(* IEC 61131-3 sources: trust-platform/examples/control/01-feedback-foundations-and-temperature-control/08-heating-valve-rate-tracking/src, 2 files *)

(* ---- Main.st ---- *)
USING Control;

(* Fraction of the raw-minus-filtered difference applied per update: alpha = dt/(Tf + dt). *)
FUNCTION FilterFraction : LREAL
VAR_INPUT
    CycleTime : LREAL;
    FilterTime : LREAL;
END_VAR
FilterFraction := CycleTime / (FilterTime + CycleTime);
END_FUNCTION

(* First-order low-pass update: yf_new = yf_old + alpha·(yr − yf_old). *)
FUNCTION FilterUpdate : LREAL
VAR_INPUT
    PreviousFilteredValue : LREAL;
    RawValue : LREAL;
    FilterFraction : LREAL;
END_VAR
FilterUpdate := PreviousFilteredValue + FilterFraction * (RawValue - PreviousFilteredValue);
END_FUNCTION

(* An interval is usable only if time has advanced and the samples can still represent the
   loop's fastest oscillation. *)
FUNCTION IntervalUsable : BOOL
VAR_INPUT
    ElapsedTime : LREAL;
    MaximumInterval : LREAL;
END_VAR
IntervalUsable := ElapsedTime > LREAL#0.0 AND ElapsedTime <= MaximumInterval;
END_FUNCTION

(* Integral correction toward the measured actuator position: I_next = I* + dt/Tt·(x − u_r). *)
FUNCTION MeasuredTrackingCorrection : LREAL
VAR_INPUT
    StemPosition : LREAL;
    Request : LREAL;
    Elapsed : LREAL;
    TrackingTime : LREAL;
END_VAR
MeasuredTrackingCorrection := Elapsed / TrackingTime * (StemPosition - Request);
END_FUNCTION

(* A reading is usable only with good source quality, inside the sensor's 0–80 °C range and with an age
   between 0 and MaximumAge. NaN fails every comparison. *)
FUNCTION ReadingUsable : BOOL
VAR_INPUT
    QualityGood : BOOL;
    Value : LREAL;
    Age : LREAL;
    MaximumAge : LREAL;
END_VAR
ReadingUsable := QualityGood AND Value >= LREAL#0.0 AND Value <= LREAL#80.0
    AND Age >= LREAL#0.0 AND Age <= MaximumAge;
END_FUNCTION

(* Weighted proportional term about the operating point T0: P = Kp·(β·(SP − T0) − (PV − T0)). *)
FUNCTION WeightedProportional : LREAL
VAR_INPUT
    ProportionalGain : LREAL;
    SetpointWeight : LREAL;
    Setpoint : LREAL;
    ProcessValue : LREAL;
    OperatingPoint : LREAL;
END_VAR
WeightedProportional := ProportionalGain
    * (SetpointWeight * (Setpoint - OperatingPoint) - (ProcessValue - OperatingPoint));
END_FUNCTION

(* Integral state that makes P + I reproduce the applied command: I = u_applied − P. *)
FUNCTION InitialIntegral : LREAL
VAR_INPUT
    AppliedOutput : LREAL;
    Proportional : LREAL;
END_VAR
InitialIntegral := AppliedOutput - Proportional;
END_FUNCTION

(* A candidate set is usable only as a whole: non-negative gains, weights in 0–1, a minimum below the
   maximum, rate limits around zero, a positive tracking time and a non-negative filter time.
   Any NaN fails its comparison and rejects the set. *)
FUNCTION ValidPidParameters : BOOL
VAR_INPUT
    Candidate : Control.PIDParameters;
    FilterTime : LREAL;
END_VAR
ValidPidParameters :=
    Candidate.ProportionalGain >= LREAL#0.0 AND Candidate.IntegralGain >= LREAL#0.0
    AND Candidate.DerivativeGain >= LREAL#0.0
    AND Candidate.ProportionalSetpointWeight >= LREAL#0.0 AND Candidate.ProportionalSetpointWeight <= LREAL#1.0
    AND Candidate.DerivativeSetpointWeight >= LREAL#0.0 AND Candidate.DerivativeSetpointWeight <= LREAL#1.0
    AND Candidate.Bias = Candidate.Bias
    AND Candidate.OutputMinimum < Candidate.OutputMaximum
    AND Candidate.RateMinimum <= LREAL#0.0 AND Candidate.RateMaximum >= LREAL#0.0
    AND Candidate.TrackingTime > LREAL#0.0
    AND FilterTime >= LREAL#0.0;
END_FUNCTION

FUNCTION SamePidParameters : BOOL
VAR_INPUT
    Left : Control.PIDParameters;
    Right : Control.PIDParameters;
END_VAR
SamePidParameters :=
    Left.ProportionalGain = Right.ProportionalGain
    AND Left.IntegralGain = Right.IntegralGain
    AND Left.DerivativeGain = Right.DerivativeGain
    AND Left.ProportionalSetpointWeight = Right.ProportionalSetpointWeight
    AND Left.DerivativeSetpointWeight = Right.DerivativeSetpointWeight
    AND Left.Bias = Right.Bias
    AND Left.OutputMinimum = Right.OutputMinimum
    AND Left.OutputMaximum = Right.OutputMaximum
    AND Left.RateMinimum = Right.RateMinimum
    AND Left.RateMaximum = Right.RateMaximum
    AND Left.TrackingTime = Right.TrackingTime
    AND Left.AntiWindup = Right.AntiWindup;
END_FUNCTION

PROGRAM Main
VAR
    Controller : Control.PID;
    (* Tune replaces this record with each candidate; the defaults are the controller commissioned
       on the electric heater in Lesson 30. *)
    Parameters : Control.PIDParameters := (
        ProportionalGain := LREAL#13.0,
        IntegralGain := LREAL#3.5,
        DerivativeGain := LREAL#0.0,
        ProportionalSetpointWeight := LREAL#0.3,
        DerivativeSetpointWeight := LREAL#0.0,
        Bias := LREAL#0.0,
        OutputMinimum := LREAL#0.0,
        OutputMaximum := LREAL#100.0,
        RateMinimum := LREAL#-10000.0,
        RateMaximum := LREAL#10000.0,
        TrackingTime := LREAL#1.0,
        AntiWindup := PIDAntiWindup#BackCalculation
    );
    ConfiguredParameters : Control.PIDParameters;
    ConfiguredFilterTimeS : LREAL := 1.0;
    ParameterRevision : DINT := 0;
    ParametersRejected : BOOL := FALSE;
    InitialState : Control.PIDInitialState;
    ObservedState : Control.PIDInitialState;
    Input : Control.PIDInput;
    (* Ready: every retained value has been set from the actual operating condition. *)
    Initialized : BOOL := FALSE;
    InitializeRequest : BOOL := FALSE;
    InitializeRequestWas : BOOL := FALSE;
    AutoMode : BOOL := FALSE;
    AutoActive : BOOL := FALSE;
    (* TRUE at start: a program that starts in Auto from preset stored values continues without a
       transfer. A real start begins uninitialized in Manual, which clears it. *)
    AutoWasActive : BOOL := TRUE;
    (* FALSE runs the untracked counterexample: Manual leaves the stored values as initialized. *)
    TrackManual : BOOL := TRUE;
    ManualOutput : LREAL := 75.0;
    (* Sensor interface: the simulated device delivers the reading with a quality flag; these three
       inputs inject faults for the lesson. *)
    SensorQualityGood : BOOL := TRUE;
    SensorFrozen : BOOL := FALSE;
    InjectedOffsetC : LREAL := 0.0;
    ReadingC : LREAL := 35.0;
    AcquisitionTimer : TON;
    AcquisitionAgeS : LREAL := 0.0;
    NewAcquisition : BOOL := FALSE;
    (* Measurement validity: a reading older than MaximumAgeS is stale; recovery needs
       FreshSamplesRequired consecutive fresh valid acquisitions after an acknowledgement. *)
    MaximumAgeS : LREAL := 0.5;
    FreshSamplesRequired : DINT := 3;
    MeasurementUsable : BOOL := FALSE;
    MeasurementFault : BOOL := FALSE;
    FaultAcknowledge : BOOL := FALSE;
    Acknowledged : BOOL := FALSE;
    RecoveryCount : DINT := 0;
    RecoveryComplete : BOOL := FALSE;
    SetpointC : LREAL := 35.0;
    TemperatureC : LREAL := 35.0;
    SafeProcessValueC : LREAL := 35.0;
    (* Requested position, bounded target and measured position: the PI request before the 0–100 %
       limits, the target sent to the valve, and the stem position the valve has reached. *)
    NominalRequestPct : LREAL := 75.0;
    ValveRequestPct : LREAL := 75.0;
    StemPositionPct : LREAL := 75.0;
    (* FALSE tracks only the bounded target: the counterexample. *)
    TrackMeasuredPosition : BOOL := TRUE;
    TrackingCorrectionPct : LREAL := 0.0;
    ErrorC : LREAL := 0.0;
    (* Reference of the weighted proportional term: the 35 °C hot operating point. *)
    OperatingPointC : LREAL := 35.0;
    (* Measurement filter: Tf = 0 bypasses it; Control Studio applies Tf with the gains. *)
    FilterTimeS : LREAL := 1.0;
    FilterAlpha : LREAL := 1.0;
    FilteredC : LREAL := 35.0;
    FilterRestart : BOOL := TRUE;
    (* Timing: the controller updates every ControllerPeriodS of measured time. *)
    IntervalTimer : TON;
    SinceLastUpdateS : LREAL := 0.0;
    ElapsedS : LREAL := 0.0;
    ControllerPeriodS : LREAL := 0.1;
    (* Longest usable interval: half the loop's 4.42 s ultimate period (Lesson 20). *)
    MaximumIntervalS : LREAL := 2.2;
    UpdateDue : BOOL := FALSE;
    TimingUsable : BOOL := FALSE;
    RejectedUpdates : DINT := 0;
    ProportionalPct : LREAL := 0.0;
    IntegralPct : LREAL := 75.0;
    PreviousRequestPct : LREAL := 75.0;
    CommandActivityPoints : LREAL := 0.0;
END_VAR

(* The water heated through the valve; the temperature measurement carries ±0.02 °C noise. *)
(* Sensor interface: every scan the device delivers a new acquisition unless it is frozen. The
   acquisition timer restarts with each new acquisition, so its elapsed time is the reading's age. *)
IF NOT SensorFrozen THEN
    ReadingC := TemperatureC + InjectedOffsetC;
    AcquisitionTimer(IN := FALSE, PT := T#1h);
    NewAcquisition := TRUE;
ELSE
    NewAcquisition := FALSE;
END_IF;
AcquisitionTimer(IN := TRUE, PT := T#1h);
AcquisitionAgeS := UDINT_TO_LREAL(DWORD_TO_UDINT(TIME_TO_DWORD(AcquisitionTimer.ET))) / LREAL#1000.0;

MeasurementUsable := ReadingUsable(QualityGood := SensorQualityGood, Value := ReadingC,
    Age := AcquisitionAgeS, MaximumAge := MaximumAgeS);
IF MeasurementUsable THEN
    SafeProcessValueC := ReadingC;
END_IF;

(* A latched fault requests a closed valve (the stem still needs time to close), stops every
   controller and filter update, and clears the Auto
   request and the manual demand, so neither can reopen the valve by itself. *)
IF NOT MeasurementUsable AND NOT MeasurementFault THEN
    MeasurementFault := TRUE;
    AutoMode := FALSE;
    ManualOutput := LREAL#0.0;
    Acknowledged := FALSE;
    RecoveryCount := 0;
END_IF;
(* Recovery: after an acknowledgement, FreshSamplesRequired consecutive new and valid acquisitions.
   A repeated old reading does not count; an invalid one restarts the count. *)
RecoveryComplete := FALSE;
IF MeasurementFault THEN
    IF FaultAcknowledge THEN
        Acknowledged := TRUE;
        FaultAcknowledge := FALSE;
        RecoveryCount := 0;
    END_IF;
    IF NOT MeasurementUsable THEN
        RecoveryCount := 0;
    ELSIF Acknowledged AND NewAcquisition THEN
        RecoveryCount := RecoveryCount + 1;
    END_IF;
    IF RecoveryCount >= FreshSamplesRequired THEN
        MeasurementFault := FALSE;
        Acknowledged := FALSE;
        RecoveryCount := 0;
        RecoveryComplete := TRUE;
    END_IF;
ELSE
    FaultAcknowledge := FALSE;
END_IF;
(* Measured time since the previous update decision, read in the scan that acquires the measurement. *)
IntervalTimer(IN := TRUE, PT := T#1h);
SinceLastUpdateS := UDINT_TO_LREAL(DWORD_TO_UDINT(TIME_TO_DWORD(IntervalTimer.ET))) / LREAL#1000.0;

(* Parameter updates: Control Studio's Apply writes the complete record and FilterTimeS at one task
   boundary. The program adopts a changed set only as a whole and only if it is valid; an invalid set
   changes nothing, and the controller keeps running on the active set. *)
IF NOT Initialized OR NOT SamePidParameters(Left := Parameters, Right := ConfiguredParameters)
        OR FilterTimeS <> ConfiguredFilterTimeS THEN
    IF ValidPidParameters(Candidate := Parameters, FilterTime := FilterTimeS) THEN
        ConfiguredParameters := Parameters;
        ConfiguredFilterTimeS := FilterTimeS;
        ParameterRevision := ParameterRevision + 1;
        ParametersRejected := FALSE;
    ELSE
        ParametersRejected := TRUE;
    END_IF;
ELSE
    ParametersRejected := FALSE;
END_IF;
Controller.Configure(Parameters := ConfiguredParameters);

(* Hot reset: the program starts with the operator's manual command at the 75 % valve position that
   holds the water at 35 °C. *)
IF NOT Initialized THEN
    ManualOutput := LREAL#75.0;
END_IF;

(* One writer for the valve request: a fault, else Manual until automatic control is active.
   Manual applies its own command and does not update the controller. *)
AutoActive := AutoMode AND Initialized AND NOT MeasurementFault
    AND ConfiguredParameters.ProportionalGain > LREAL#0.0 AND ConfiguredParameters.IntegralGain > LREAL#0.0;
IF MeasurementFault THEN
    ValveRequestPct := LREAL#0.0;
ELSIF NOT AutoActive THEN
    ValveRequestPct := LIMIT(MN := LREAL#0.0, IN := ManualOutput, MX := LREAL#100.0);
END_IF;

(* Initialization sets every retained value from the actual operating condition: at startup and
   once per rising edge of InitializeRequest, only while Manual owns the valve and the data is valid. *)
IF (NOT Initialized OR (InitializeRequest AND NOT InitializeRequestWas) OR RecoveryComplete)
        AND NOT AutoActive AND NOT MeasurementFault AND MeasurementUsable THEN
    IF NOT Initialized AND NOT AutoMode THEN
        SetpointC := SafeProcessValueC;
    END_IF;
    FilteredC := SafeProcessValueC;
    InitialState.Setpoint := SetpointC;
    InitialState.ProcessValue := FilteredC;
    InitialState.NominalOutput := ValveRequestPct;
    InitialState.SaturatedOutput := ValveRequestPct;
    InitialState.SetpointRate := LREAL#0.0;
    InitialState.ProcessValueRate := LREAL#0.0;
    InitialState.FeedForward := LREAL#0.0;
    Controller.Initialize(State := InitialState);
    ProportionalPct := WeightedProportional(ProportionalGain := ConfiguredParameters.ProportionalGain,
        SetpointWeight := ConfiguredParameters.ProportionalSetpointWeight, Setpoint := SetpointC,
        ProcessValue := FilteredC, OperatingPoint := OperatingPointC);
    IntegralPct := InitialIntegral(AppliedOutput := ValveRequestPct, Proportional := ProportionalPct);
    NominalRequestPct := ValveRequestPct;
    Initialized := TRUE;
END_IF;
InitializeRequestWas := InitializeRequest;

(* Manual keeps the timing baseline current every scan, so the first automatic update integrates
   one scan, not the time spent in Manual. Auto updates every ControllerPeriodS. *)
UpdateDue := NOT AutoActive OR NOT AutoWasActive
    OR SinceLastUpdateS >= ControllerPeriodS - LREAL#0.001;
IF UpdateDue THEN
    ElapsedS := SinceLastUpdateS;
    TimingUsable := IntervalUsable(ElapsedTime := ElapsedS, MaximumInterval := MaximumIntervalS);
    IntervalTimer(IN := FALSE, PT := T#1h);
    IntervalTimer(IN := TRUE, PT := T#1h);
END_IF;
IF UpdateDue AND NOT TimingUsable THEN
    (* No state is updated over an unusable interval: the command is held, and the next
       accepted update restarts the filter from the fresh measurement. *)
    IF AutoActive THEN
        RejectedUpdates := RejectedUpdates + 1;
    END_IF;
    FilterRestart := TRUE;
ELSIF UpdateDue AND NOT MeasurementFault THEN
    (* The filter runs in Auto; in Manual, on the transfer scan and after a restart it takes the fresh measurement. *)
    IF AutoActive AND AutoWasActive AND NOT FilterRestart THEN
        FilterAlpha := FilterFraction(CycleTime := ElapsedS, FilterTime := ConfiguredFilterTimeS);
        FilteredC := FilterUpdate(PreviousFilteredValue := FilteredC, RawValue := SafeProcessValueC, FilterFraction := FilterAlpha);
    ELSE
        FilteredC := SafeProcessValueC;
    END_IF;
    FilterRestart := FALSE;
    Input.Setpoint := SetpointC;
    Input.ProcessValue := FilteredC;
    Input.CycleTime := ElapsedS;
    Input.FeedForward := LREAL#0.0;
    Input.TrackingOutput := ValveRequestPct;
    Input.ManualOutput := ValveRequestPct;
    ErrorC := SetpointC - FilteredC;
    IF AutoActive AND (AutoWasActive OR NOT TrackManual) THEN
        (* Ordinary PI update. *)
        Input.Mode := PIDMode#Auto;
        ValveRequestPct := Controller.Update(Input := Input);
        AutoWasActive := TRUE;
        (* Measured-position tracking: move the integral toward the stem position the valve has
           reached, with the controller's tracking time. *)
        IF TrackMeasuredPosition AND StemPositionPct >= LREAL#0.0 AND StemPositionPct <= LREAL#100.0 THEN
            TrackingCorrectionPct := MeasuredTrackingCorrection(StemPosition := StemPositionPct,
                Request := ValveRequestPct, Elapsed := ElapsedS, TrackingTime := ConfiguredParameters.TrackingTime);
            ObservedState := Controller.GetState();
            ObservedState.NominalOutput := ObservedState.NominalOutput + TrackingCorrectionPct;
            Controller.Initialize(State := ObservedState);
        ELSE
            TrackingCorrectionPct := LREAL#0.0;
        END_IF;
    ELSIF TrackManual THEN
        (* Tracking: in Manual and on the transfer scan, the stored values follow the applied command,
           the setpoint and the measurement, so I = u_a − P. The command stays u_a: no integral step. *)
        Input.Mode := PIDMode#Manual;
        ValveRequestPct := Controller.Update(Input := Input);
        AutoWasActive := AutoActive;
    END_IF;

    (* Diagnostics come from the actual controller state; the PI equations live in Control.PID. *)
    ObservedState := Controller.GetState();
    NominalRequestPct := ObservedState.NominalOutput;
    ProportionalPct := WeightedProportional(ProportionalGain := ConfiguredParameters.ProportionalGain,
        SetpointWeight := ConfiguredParameters.ProportionalSetpointWeight, Setpoint := SetpointC,
        ProcessValue := FilteredC, OperatingPoint := OperatingPointC);
    IntegralPct := NominalRequestPct - ProportionalPct;
END_IF;
IF NOT AutoActive THEN
    AutoWasActive := FALSE;
END_IF;
(* Command activity adds every applied-command movement, starting from the 75 % holding command. *)
CommandActivityPoints := CommandActivityPoints + ABS(ValveRequestPct - PreviousRequestPct);
PreviousRequestPct := ValveRequestPct;

END_PROGRAM

CONFIGURATION Config
RESOURCE Res ON PLC
    TASK MainTask(INTERVAL := T#100ms, PRIORITY := 1);
    PROGRAM P1 WITH MainTask : Main;
END_RESOURCE
VAR_CONFIG
    P1.MeasurementFault AT %MX96.3 : BOOL;
    P1.MeasurementUsable AT %MX96.2 : BOOL;
    P1.ValveRequestPct AT %QL0 : LREAL;
    P1.TemperatureC AT %IL8 : LREAL;
    P1.StemPositionPct AT %IL16 : LREAL;
    P1.SetpointC AT %ML0 : LREAL;
    P1.IntegralPct AT %ML16 : LREAL;
    P1.NominalRequestPct AT %ML32 : LREAL;
    P1.ProportionalPct AT %ML56 : LREAL;
    P1.CommandActivityPoints AT %ML64 : LREAL;
    P1.ManualOutput AT %ML72 : LREAL;
END_VAR
END_CONFIGURATION

(* ---- tests.st ---- *)
(* @trustlsp:runtime-ignore — run these assertions with trust-dev test;
   they are not scheduled PLC instances in the lesson simulator. *)

TEST_PROGRAM TrackingMovesTheIntegralTowardTheStem
(* Stem at 75 %, request 80.1 %, dt = 0.1 s, Tt = 1 s: the integral moves by -0.51 point. *)
ASSERT_NEAR(EXPECTED := LREAL#-0.51, ACTUAL := MeasuredTrackingCorrection(StemPosition := LREAL#75.0,
    Request := LREAL#80.1, Elapsed := LREAL#0.1, TrackingTime := LREAL#1.0), DELTA := LREAL#1.0e-9);
(* A stem that has reached the request needs no correction. *)
ASSERT_NEAR(EXPECTED := LREAL#0.0, ACTUAL := MeasuredTrackingCorrection(StemPosition := LREAL#80.0,
    Request := LREAL#80.0, Elapsed := LREAL#0.1, TrackingTime := LREAL#1.0), DELTA := LREAL#1.0e-12);
END_TEST_PROGRAM

TEST_PROGRAM RateLimitSetsTheTravelTime
VAR
    Seconds : LREAL;
END_VAR
(* At 0.5 % per second, 75 → 85 % takes 10 points / 0.5 %/s = 20 s. *)
Seconds := (LREAL#85.0 - LREAL#75.0) / LREAL#0.5;
ASSERT_NEAR(EXPECTED := LREAL#20.0, ACTUAL := Seconds, DELTA := LREAL#1.0e-12);
END_TEST_PROGRAM
